Fanuc KAREL source: KC00016.KL

PROGRAM KC00016
%NOLOCKGROUP
%ENVIRONMENT MULTI
VAR
  I: INTEGER
  J: INTEGER
  K: INTEGER
  R: REAL
  B: BOOLEAN
  S: STRING[80]
  T: STRING[80]
  P: PATH
  Q: PATH
  AI: ARRAY[8] OF INTEGER
  AB: ARRAY[244] OF BYTE
BEGIN
  POST_SEMA(I)
END KC00016
